TYPE ST_AnalogSignal :
STRUCT
	//analog signal
	nIn_RawSignal	:	UINT		;
	rOut_Converted	:	REAL	;
	
	//analog signal settings
	rRawMax	:	REAL:=32767	;
	rRawMin	:	REAL:=0		;
	rOutMax	:	REAL:=100	;
	rOutMin	:	REAL:=10 	;
	//not usable 
	rRawZeroPointOffset	:	REAL:=100;//offset foranalog signal //?
	rRawMaxPointOffset	:	INT:=100;//?
END_STRUCT
END_TYPE

(* stored: Version 1.1.0.1, ProductVersion 3.1.4024.12
   DUT ST_AnalogSignal: Id {d8cd7068-f878-40c3-8d17-e3dd45112344} *)
